(* IEC 61131-3 sources: Mori.EscaFlow/tests/Conformance/golden/logix, 9 files *)

(* ---- aoi.st ---- *)
FUNCTION_BLOCK Motor
VAR_INPUT
    EnableIn : BOOL;
    Cmd : BOOL; (* run command *)
    Speed : REAL;
    Delay : DINT := 500;
END_VAR
VAR_OUTPUT
    EnableOut : BOOL;
    Running : BOOL;
    Fault : BOOL;
END_VAR
VAR_IN_OUT
    Data : MotorData;
END_VAR
VAR RETAIN
    T1 : TIMER;
    Count : DINT;
    Prev : BOOL;
END_VAR

VAR_TEMP
    _rc1 : BOOL;
END_VAR
T1(IN := Cmd); (* TON/logix *)
Running := Cmd AND T1.DN;
_rc1 := R_EDGE(Cmd, Prev);
IF _rc1 THEN
    Data.Starts := Data.Starts + 1;
END_IF;
IF _rc1 THEN
    Count := Count + 1;
END_IF;
Fault := Running AND Speed > 100.0;

ACTION Prescan
    Running := 0;
    Count := 0;
END_ACTION

ACTION Postscan (* hook: postscan *)
    Running := 0;
END_ACTION

ACTION EnableInFalse (* hook: enableFalse *)
    Running := 0;
    Fault := 0;
END_ACTION

ACTION Init (* hook: init *)
    T1(IN := FALSE); (* TON/logix, mode: prescan *)
    Running := FALSE;
    Prev := TRUE;
    Fault := FALSE;
    Prescan();
END_ACTION
END_FUNCTION_BLOCK

PROGRAM P

Main();

ACTION Main
    M1(EN := Start, Cmd := Start, Speed := Spd, Data := MD1, Running => Run1); (* Motor *)
    Text();
END_ACTION

ACTION Text
    M2(Cmd := Start, Speed := Spd, Data := MD2, Running => Run2); (* Motor *)
    M2.Delay := 250;
    Run2 := M2.Running AND NOT M2.Fault;
END_ACTION

ACTION Prescan (* hook: init *)
    M1(Data := MD1); (* Motor, mode: prescan *)
    M2(Data := MD2); (* Motor, mode: prescan *)
END_ACTION
END_PROGRAM

(* ---- fbd.st ---- *)
FUNCTION_BLOCK Blink
VAR_INPUT
    EnableIn : BOOL;
    Rate : DINT;
    Reset : BOOL;
END_VAR
VAR_OUTPUT
    EnableOut : BOOL;
    Out : BOOL;
END_VAR
VAR_IN_OUT
    Data : DINT;
END_VAR
VAR RETAIN
    T1 : TIMER;
END_VAR

T1.PRE := Rate;
Out := T1.DN AND NOT Reset;
Data := Data + 1;

ACTION Init (* hook: init *)
END_ACTION
END_FUNCTION_BLOCK

PROGRAM P
VAR RETAIN
    InA : DINT;
    OutA : DINT;
END_VAR

Main();

ACTION Main
    VAR_TEMP
        _f1 : REAL;
    END_VAR
    TONR_01.TimerEnable := In1;
    TONR_01.PRE := Preset;
    TONR_01.Reset := Blink_01.Out;
    TONR(TONR_01); (* logix *)
    Out1 := TONR_01.DN;
    Blink_01.Rate := Preset;
    Blink_01.Reset := TONR_01.DN;
    Blink_01(Data := Counter); (* Blink *)
    Out2 := Blink_01.Out;
    _f1 := Val + 1.5;
    SumOut := _f1;
    InA := Preset;
    Sub();
    RetVal := OutA;
END_ACTION

ACTION Sub
    OutA := InA + 1;
    RETURN;
END_ACTION

ACTION Prescan (* hook: init *)
    TONR(TONR_01); (* logix *)
    Blink_01(Data := Counter); (* Blink, mode: prescan *)
END_ACTION
END_PROGRAM

(* ---- ladder.st ---- *)
FUNCTION_BLOCK Blink
VAR_INPUT
    EnableIn : BOOL;
    Rate : DINT;
END_VAR
VAR_OUTPUT
    EnableOut : BOOL;
    Out : BOOL;
END_VAR
VAR RETAIN
    T1 : TIMER;
END_VAR

VAR_TEMP
    _rc1 : BOOL;
END_VAR
_rc1 := NOT T1.DN;
T1(IN := _rc1); (* TON/logix *)
Out := NOT T1.DN AND T1.DN;

ACTION Init (* hook: init *)
    T1(IN := FALSE); (* TON/logix, mode: prescan *)
    Out := FALSE;
END_ACTION
END_FUNCTION_BLOCK

PROGRAM P
VAR RETAIN
    InA : DINT;
    InB : DINT;
    OutA : DINT;
END_VAR

Main();

ACTION Main
    VAR_TEMP
        _rc1 : BOOL;
        _rc2 : BOOL;
        _rc3 : BOOL;
        _mcr1 : BOOL;
        _rc4 : BOOL;
    END_VAR
    _rc1 := A AND NOT B;
    Out1 := _rc1;
    IF _rc1 THEN
        Out2 := TRUE;
    END_IF;
    IF _rc1 THEN
        Bits.3 := FALSE;
    END_IF;
    _rc2 := R_EDGE(A, Bits.0);
    Pulse := R_EDGE(_rc2, Bits.1);
    C := F_EDGE(_rc2, Bits.2);
    Out1 := X = Y AND X <> 1 AND X > 2 AND Y >= X AND Z < X AND Z <= Y AND X + Y > Z AND (0 <= 10 AND (0 <= X AND X <= 10) OR 0 > 10 AND (X >= 0 OR X <= 10)) AND (Bits AND 16#FF) = (Y AND 16#FF);
    T1(IN := A); (* TON/logix *)
    T2(IN := A); (* TOF/logix *)
    T3(IN := A); (* TONR/logix *)
    C1(CU := A); (* CTU/logix *)
    C2(CD := A); (* CTD/logix *)
    _rc3 := A AND B;
    IF _rc3 THEN
        T3.ACC := 0;
        T3.EN := FALSE;
        T3.TT := FALSE;
        T3.DN := FALSE;
    END_IF;
    IF _rc3 THEN
        C1.ACC := 0;
        C1.CU := FALSE;
        C1.CD := FALSE;
        C1.DN := FALSE;
        C1.OV := FALSE;
        C1.UN := FALSE;
    END_IF;
    IF A THEN
        Y := X;
    END_IF;
    IF A THEN
        Z := 0;
    END_IF;
    IF A THEN
        Z := X + Y;
    END_IF;
    IF A THEN
        Z := X - 1;
    END_IF;
    IF A THEN
        Z := X * 2;
    END_IF;
    IF A THEN
        Z := X / Y;
    END_IF;
    IF A THEN
        Z := X MOD 3;
    END_IF;
    IF A THEN
        Bits := X AND Y;
    END_IF;
    IF A THEN
        Bits := X OR 16#F;
    END_IF;
    IF A THEN
        Bits := Bits XOR Y;
    END_IF;
    IF A THEN
        Y := NOT X;
    END_IF;
    IF A THEN
        Z := -X;
    END_IF;
    IF A THEN
        R := ABS(R);
    END_IF;
    IF A THEN
        R := SQRT(R);
    END_IF;
    IF A THEN
        Z := TO_DINT#roundEven((X + Y) * 2 - R);
    END_IF;
    IF B THEN
        COPY(Src[0], Dst[0], 10); (* bytes *)
    END_IF;
    IF B THEN
        COPY_ATOMIC(Src[0], Dst[0], 10); (* bytes *)
    END_IF;
    IF B THEN
        FILL(0, Dst[0], 10);
    END_IF;
    IF A THEN
        InA := X;
        InB := Y;
        Sub();
        Z := OutA;
    END_IF;
    IF C THEN
        JMP Skip;
    END_IF;
    Out2 := A AND (B OR C AND (NOT A OR Out1) OR X = Y);
    Skip:
    _mcr1 := A;
    _rc4 := _mcr1 AND B;
    Out1 := _rc4;
    T1(IN := _rc4); (* TON/logix *)
    Out1 := FALSE;
    IF A THEN
        GSV(WallClockTime, , DateTime, Clock[0]); (* logix *)
    END_IF;
    IF A THEN
        SSV(Program, P, DisableFlag, X); (* logix *)
    END_IF;
    (* EN := A *) MSG(Msg1); (* logix *)
    Blk(EN := A, Rate := 250, Out => Out2); (* Blink *)
    IF A THEN
        Y := BIT_FIELD_DISTRIBUTE(X, 0, Y, 8, 4);
    END_IF;
    IF A THEN
        Bits := MASKED_MOVE(X, 16#FF00, Bits);
    END_IF;
    IF A THEN
        Y := SWAP_BYTES(X, REVERSE);
    END_IF;
    IF A THEN
        S3 := CONCAT(S1, S2);
    END_IF;
    IF A THEN
        S2 := MID(S1, 3, 1);
    END_IF;
    IF A THEN
        Idx := FIND(S1, S2, 1);
    END_IF;
    IF A THEN
        FOR Idx := 0 TO 9 BY 1 DO
            Loop();
        END_FOR;
    END_IF;
    IF B THEN
        RETURN;
    END_IF;
END_ACTION

ACTION Sub
    OutA := InA + InB;
    RETURN;
END_ACTION

ACTION Loop
    Dst[Idx] := Idx;
    IF Dst[Idx] = 5 THEN
        BRK(); (* logix *)
    END_IF;
END_ACTION

ACTION Prescan (* hook: init *)
    Out1 := FALSE;
    Bits.0 := TRUE;
    Pulse := FALSE;
    Bits.1 := TRUE;
    C := FALSE;
    Bits.2 := TRUE;
    Out1 := FALSE;
    T1(IN := FALSE); (* TON/logix, mode: prescan *)
    T2(IN := FALSE); (* TOF/logix, mode: prescan *)
    T3(IN := FALSE); (* TONR/logix, mode: prescan *)
    C1(CU := FALSE); (* CTU/logix, mode: prescan *)
    C2(CD := FALSE); (* CTD/logix, mode: prescan *)
    Out2 := FALSE;
    Out1 := FALSE;
    T1(IN := FALSE); (* TON/logix, mode: prescan *)
    Out1 := FALSE;
    MSG(Msg1); (* logix *)
    Blk(); (* Blink, mode: prescan *)
END_ACTION
END_PROGRAM

(* ---- st.st ---- *)
FUNCTION_BLOCK Blink
VAR_INPUT
    EnableIn : BOOL;
    Rate : DINT;
END_VAR
VAR_OUTPUT
    EnableOut : BOOL;
    Out : BOOL;
END_VAR
VAR RETAIN
    T1 : TIMER;
END_VAR

T1.PRE := Rate;
TONR(T1); (* logix *)
Out := T1.DN;

ACTION Init (* hook: init *)
    TONR(T1); (* logix *)
END_ACTION
END_FUNCTION_BLOCK

PROGRAM P
VAR RETAIN
    InA : DINT;
    OutA : DINT;
END_VAR

Main();

ACTION Main
    D := TO_DINT#roundEven(R * 2.0);
    S := TO_SINT#wrap(D + 1);
    R := TO_REAL#roundEven(L);
    L := D / 3;
    IF D > 10 AND NOT Flag THEN
        D := 0;
    ELSIF D < 0 OR Flag THEN
        D := 10;
    ELSE
        D := D + 1;
    END_IF;
    CASE D OF
        1:
            Flag := 1;
        2..5, 8:
            Flag := 0;
        ELSE
            Flag := D.0;
    END_CASE;
    FOR I := 0 TO 4 BY 1 DO
        Arr[I] := I * 2;
        IF Arr[I] > 6 THEN
            EXIT;
        END_IF;
    END_FOR;
    WHILE I > 0 DO
        I := I - 1;
    END_WHILE;
    REPEAT
        I := I + 1;
    UNTIL I >= 3
    END_REPEAT;
    R := ABS(R) + SQRT(R) - SIN(R);
    D := TRUNC(R);
    Word.[I] := 1;
    Flag := Word.[D];
    D := Str.LEN;
    Str.DATA[0] := TO_SINT#wrap(65);
    Str2 := Str;
    IF TRUE THEN
        InA := D;
        Sub();
        Word := OutA;
    END_IF;
    Blk(Rate := 100, Out => Flag); (* Blink *)
    Flag := D >= 5 XOR Flag;
END_ACTION

ACTION Sub
    OutA := InA * 2;
    RETURN;
END_ACTION

ACTION Prescan (* hook: init *)
    Blk(); (* Blink, mode: prescan *)
END_ACTION
END_PROGRAM

(* ---- messages.st ---- *)
PROGRAM P
VAR RETAIN
    State : DINT;
END_VAR

Main();

ACTION Main
    VAR_TEMP
        _rc1 : BOOL;
        _rc2 : BOOL;
        _rc3 : BOOL;
        _rc4 : BOOL;
        _rc5 : BOOL;
    END_VAR
    (* EN := Trigger AND NOT Read_Remote.EN *) MSG(Read_Remote); (* logix *)
    _rc1 := State = 0;
    IF _rc1 THEN
        MsgData.Create_Source.Type := 1;
    END_IF;
    IF _rc1 THEN
        MsgData.Create_Source.Addr.Family := TO_INT#wrap(2);
    END_IF;
    IF _rc1 THEN
        MsgData.Create_Source.Addr.Port := TO_INT#wrap(5000);
    END_IF;
    (* EN := _rc1 *) MSG(SKT_Create); (* logix *)
    IF SKT_Create.DN THEN
        SKT_Open.Instance := MsgData.Instance;
    END_IF;
    IF SKT_Create.DN THEN
        SKT_Write.Instance := MsgData.Instance;
    END_IF;
    IF SKT_Create.DN THEN
        SKT_Read.Instance := MsgData.Instance;
    END_IF;
    IF SKT_Create.DN THEN
        SKT_Delete.Instance := MsgData.Instance;
    END_IF;
    IF SKT_Create.DN THEN
        State := 1;
    END_IF;
    _rc2 := State = 1;
    (* EN := _rc2 *) MSG(SKT_Open); (* logix *)
    IF State = 1 AND SKT_Open.DN THEN
        State := 2;
    END_IF;
    _rc3 := State = 2;
    (* EN := _rc3 *) MSG(SKT_Write); (* logix *)
    IF State = 2 AND SKT_Write.DN THEN
        State := 3;
    END_IF;
    _rc4 := State = 3;
    (* EN := _rc4 *) MSG(SKT_Read); (* logix *)
    IF State = 3 AND SKT_Read.DN THEN
        State := 4;
    END_IF;
    _rc5 := State = 4;
    (* EN := _rc5 *) MSG(SKT_Delete); (* logix *)
    IF State = 4 AND SKT_Delete.DN THEN
        State := 0;
    END_IF;
    (* EN := Trigger *) MSG(Get_Identity); (* logix *)
    IF Trigger THEN
        ProdCount := ConsCount;
    END_IF;
END_ACTION

ACTION Prescan (* hook: init *)
    MSG(Read_Remote); (* logix *)
    MSG(SKT_Create); (* logix *)
    MSG(SKT_Open); (* logix *)
    MSG(SKT_Write); (* logix *)
    MSG(SKT_Read); (* logix *)
    MSG(SKT_Delete); (* logix *)
    MSG(Get_Identity); (* logix *)
END_ACTION
END_PROGRAM

(* ---- modules.st ---- *)
PROGRAM P

Main();

ACTION Main
    Flag := DI:I.Data.4 AND NOT DI:I.Fault.0;
    ENet:O.Data[0] := Word;
    Word := ENet:I.Data[1] + DI:I.Data;
    Cfg := Turck:C.Channel_Mode_Port1;
    Byte0 := Turck:I.Data[0];
    Flag := Turck:I.ConnectionFaulted OR ENet:I.Data[1].0 OR DI:I.Data.4;
    DI:O.Data.0 := Flag;
END_ACTION

ACTION Prescan (* hook: init *)
END_ACTION
END_PROGRAM

(* ---- sfc.st ---- *)
PROGRAM P
VAR RETAIN
    Step_000 : SFC_STEP;
    Step_001 : SFC_STEP;
    Step_002 : SFC_STEP;
    Step_003 : SFC_STEP;
    Step_004 : SFC_STEP;
    Tran_000 : BOOL;
    Tran_001 : BOOL;
    Tran_002 : BOOL;
    Tran_003 : BOOL;
    Action_000 : SFC_ACTION;
    Action_001 : SFC_ACTION;
    Action_002 : SFC_ACTION;
    Action_003 : SFC_ACTION;
    Action_004 : SFC_ACTION;
    Action_005 : SFC_ACTION;
    Action_006 : SFC_ACTION;
    Action_007 : SFC_ACTION;
    Action_008 : SFC_ACTION;
    Stop_000 : SFC_STOP;
END_VAR

Main();

ACTION Main
END_ACTION

ACTION Prescan (* hook: init *)
END_ACTION
END_PROGRAM

(* ---- tasks.st ---- *)
PROGRAM P1
VAR RETAIN
    Local1 : DINT;
END_VAR

Main();

ACTION Main
    Counter := Counter + 1;
END_ACTION

ACTION Fault
    Local1 := 0;
END_ACTION

ACTION Prescan (* hook: init *)
END_ACTION
END_PROGRAM

PROGRAM P2

Main();

ACTION Main
    Counter := 0;
END_ACTION

ACTION Prescan (* hook: init *)
END_ACTION
END_PROGRAM

PROGRAM P3

Main();

ACTION Main
    Counter := Counter - 1;
END_ACTION

ACTION Prescan (* hook: init *)
END_ACTION
END_PROGRAM

PROGRAM P4

Main();

ACTION Main
    Counter := Cons;
END_ACTION

ACTION Prescan (* hook: init *)
END_ACTION
END_PROGRAM

PROGRAM Folder

ACTION Prescan (* hook: init *)
END_ACTION
END_PROGRAM

(* ---- types.st ---- *)
PROGRAM P
VAR RETAIN
    Local : Outer;
END_VAR

Main();

ACTION Main
    O.In.Value := O.In.Value + 1.0;
    IF O.In.Bit1 AND Word.5 AND O.In.Flags[3] THEN
        Matrix[1, 2] := O.Count;
    END_IF;
    O.Items[1].Words[2] := Matrix[0, 1] + Local.Items[0].Words[3];
    O.Name := Label;
    O.Count := O.Short.LEN + O.Timer.PRE + O.Counter.ACC + O.Control.POS;
END_ACTION

ACTION Prescan (* hook: init *)
END_ACTION
END_PROGRAM
